// Position nommée (docs/06 § 2)
{attribute 'pack_mode' := '1'}
TYPE ST_NamedPos :
STRUCT
    stPos : ST_Position;
    fApproach : LREAL;
    bTaught : BOOL;
END_STRUCT
END_TYPE

(* stored: Version 1.1.0.1, ProductVersion 3.1.4024.12
   DUT ST_NamedPos: Id {7e067a51-5fd7-5e5e-a690-e062db81f5a4} *)
